TYPE "DT_DIGITAL_INPUT_HPU_PUMPS"
VERSION : 0.1
   STRUCT
      PUMP_1_THERMAL_PROT { S7_SetPoint := 'False'} : "DT_STATUS_SOLO" := ((FALSE, 1, 256), (32000, 32000, 32000), (0, 0, 0), (FALSE, FALSE, 0));
      PUMP_1_REMOTE_SWITCH { S7_SetPoint := 'False'} : "DT_STATUS_SOLO" := ((FALSE, 1, 257), (32000, 32000, 32000), (0, 0, 0), (FALSE, FALSE, 0));
      PUMP_1_TRIPPED { S7_SetPoint := 'False'} : "DT_STATUS_SOLO" := ((FALSE, 1, 258), (32000, 32000, 32000), (0, 0, 0), (FALSE, FALSE, 0));
      PUMP_1_MCB_ON { S7_SetPoint := 'False'} : "DT_STATUS_SOLO" := ((FALSE, 1, 259), (32000, 32000, 32000), (0, 3, 4), (FALSE, FALSE, 0));
      PUMP_1_CONT_ON { S7_SetPoint := 'False'} : "DT_STATUS_SOLO" := ((FALSE, 1, 260), (32000, 32000, 32000), (0, 1, 4), (FALSE, FALSE, 0));
      PUMP_2_THERMAL_PROT { S7_SetPoint := 'False'} : "DT_STATUS_SOLO" := ((FALSE, 1, 261), (32000, 32000, 32000), (0, 0, 0), (FALSE, FALSE, 0));
      PUMP_2_REMOTE_SWITCH { S7_SetPoint := 'False'} : "DT_STATUS_SOLO" := ((FALSE, 1, 262), (32000, 32000, 32000), (0, 0, 0), (FALSE, FALSE, 0));
      PUMP_2_TRIPPED { S7_SetPoint := 'False'} : "DT_STATUS_SOLO" := ((FALSE, 1, 263), (32000, 32000, 32000), (0, 0, 0), (FALSE, FALSE, 0));
      PUMP_2_ON { S7_SetPoint := 'False'} : "DT_STATUS_SOLO" := ((FALSE, 1, 264), (32000, 32000, 32000), (0, 3, 4), (FALSE, FALSE, 0));
      PUMP_2_CONT_ON { S7_SetPoint := 'False'} : "DT_STATUS_SOLO" := ((FALSE, 1, 265), (32000, 32000, 32000), (0, 1, 4), (FALSE, FALSE, 0));
      PUMP_DC_THERMAL_PROT { S7_SetPoint := 'False'} : "DT_STATUS_SOLO" := ((FALSE, 1, 266), (32000, 32000, 32000), (0, 1, 3), (FALSE, FALSE, 0));
      PUMP_DC_REMOTE_SWITCH { S7_SetPoint := 'False'} : "DT_STATUS_SOLO" := ((FALSE, 1, 267), (32000, 32000, 32000), (0, 0, 0), (FALSE, FALSE, 0));
      PUMP_DC_TRIPPED { S7_SetPoint := 'False'} : "DT_STATUS_SOLO" := ((FALSE, 1, 268), (32000, 32000, 32000), (0, 0, 0), (FALSE, FALSE, 0));
      PUMP_DC_MCB_ON { S7_SetPoint := 'False'} : "DT_STATUS_SOLO" := ((FALSE, 1, 269), (32000, 32000, 32000), (0, 0, 0), (FALSE, FALSE, 0));
      PUMP_DC_CONT_ON { S7_SetPoint := 'False'} : "DT_STATUS_SOLO" := ((FALSE, 1, 270), (32000, 32000, 32000), (0, 0, 0), (FALSE, FALSE, 0));
      SPARE_271 { S7_SetPoint := 'False'} : "DT_STATUS_SOLO" := ((FALSE, 1, 271), (32000, 32000, 32000), (0, 0, 0), (FALSE, FALSE, 0));
      SPARE_272 { S7_SetPoint := 'False'} : "DT_STATUS_SOLO" := ((FALSE, 1, 272), (32000, 32000, 32000), (0, 0, 0), (FALSE, FALSE, 0));
      SPARE_273 { S7_SetPoint := 'False'} : "DT_STATUS_SOLO" := ((FALSE, 1, 273), (32000, 32000, 32000), (0, 0, 0), (FALSE, FALSE, 0));
      SPARE_274 { S7_SetPoint := 'False'} : "DT_STATUS_SOLO" := ((FALSE, 1, 274), (32000, 32000, 32000), (0, 0, 0), (FALSE, FALSE, 0));
      SPARE_275 { S7_SetPoint := 'False'} : "DT_STATUS_SOLO" := ((FALSE, 1, 275), (32000, 32000, 32000), (0, 0, 0), (FALSE, FALSE, 0));
      SPARE_276 { S7_SetPoint := 'False'} : "DT_STATUS_SOLO" := ((FALSE, 1, 276), (32000, 32000, 32000), (0, 0, 0), (FALSE, FALSE, 0));
      SPARE_277 { S7_SetPoint := 'False'} : "DT_STATUS_SOLO" := ((FALSE, 1, 277), (32000, 32000, 32000), (0, 0, 0), (FALSE, FALSE, 0));
      SPARE_278 { S7_SetPoint := 'False'} : "DT_STATUS_SOLO" := ((FALSE, 1, 278), (32000, 32000, 32000), (0, 0, 0), (FALSE, FALSE, 0));
      SPARE_279 { S7_SetPoint := 'False'} : "DT_STATUS_SOLO" := ((FALSE, 1, 279), (32000, 32000, 32000), (0, 0, 0), (FALSE, FALSE, 0));
      SPARE_280 { S7_SetPoint := 'False'} : "DT_STATUS_SOLO" := ((FALSE, 1, 280), (32000, 32000, 32000), (0, 0, 0), (FALSE, FALSE, 0));
      SPARE_281 { S7_SetPoint := 'False'} : "DT_STATUS_SOLO" := ((FALSE, 1, 281), (32000, 32000, 32000), (0, 0, 0), (FALSE, FALSE, 0));
      SPARE_282 { S7_SetPoint := 'False'} : "DT_STATUS_SOLO" := ((FALSE, 1, 282), (32000, 32000, 32000), (0, 0, 0), (FALSE, FALSE, 0));
      SPARE_283 { S7_SetPoint := 'False'} : "DT_STATUS_SOLO" := ((FALSE, 1, 283), (32000, 32000, 32000), (0, 0, 0), (FALSE, FALSE, 0));
      SPARE_284 { S7_SetPoint := 'False'} : "DT_STATUS_SOLO" := ((FALSE, 1, 284), (32000, 32000, 32000), (0, 0, 0), (FALSE, FALSE, 0));
      SPARE_285 { S7_SetPoint := 'False'} : "DT_STATUS_SOLO" := ((FALSE, 1, 285), (32000, 32000, 32000), (0, 0, 0), (FALSE, FALSE, 0));
      SPARE_286 { S7_SetPoint := 'False'} : "DT_STATUS_SOLO" := ((FALSE, 1, 286), (32000, 32000, 32000), (0, 0, 0), (FALSE, FALSE, 0));
      SPARE_287 { S7_SetPoint := 'False'} : "DT_STATUS_SOLO" := ((FALSE, 1, 287), (32000, 32000, 32000), (0, 0, 0), (FALSE, FALSE, 0));
   END_STRUCT;

END_TYPE

